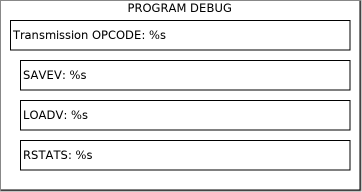
VISUALIZATION PROGRAM_STATUS  // 362x192
    Rectangle (0,0 360x190), "PROGRAM DEBUG"
    Rectangle (10,20 340x30), "Transmission OPCODE: %s", text variable: MAIN.OPCODE
    Rectangle (20,60 330x30), "SAVEV: %s", text variable: MAIN.SAVEV.ESERVER.eState
    Rectangle (20,100 330x30), "LOADV: %s", text variable: MAIN.LOADV.eState
    Rectangle (20,140 330x30), "RSTATS: %s", text variable: MAIN.RSTATS.ESERVER.eState
END_VISUALIZATION

(* stored: Version 1.1.0.1, ProductVersion 3.1.4024.16
   Visu PROGRAM_STATUS: Id {e728867c-3bb4-406b-9910-3afe4a1f041e} *)
